Fanuc KAREL source: kt00374.KL

-- PROVISIONAL review KL for V1013-1; original PC SHA256 1d1ada5c01374feee69af134d6d6749db33f4e75e4cc2827b566695011ad0318
-- Incomplete behavior may be omitted. Consult companion uncertainty JSON. Do not deploy.
PROGRAM KT00374
%NOLOCKGROUP
VAR
  S1 : STRING[80]
  S2 : STRING[80]
  OUT : BOOLEAN
BEGIN
  -- UNRESOLVED_PC offsets 5-14; opcodes 3F,75
  -- UNRESOLVED_PC offsets 19-28; opcodes 3F,75
  -- UNRESOLVED_PC offsets 33-42; opcodes 3F,75
  -- UNRESOLVED_PC offsets 47-56; opcodes 3F,75
  -- UNRESOLVED_PC offsets 61-80; opcodes 73,73,86,23
  -- UNRESOLVED_PC offsets 85-89; opcodes 7F
END KT00374
